// TIA Portal V20 export
Screen "OP01Pop-up_PRBWork"  274x350
  ScreenItem "Text field TG Status" at 1,0 size 273x47  Type=HmiTextBox
  ScreenItem "Cancel Mode" at 195,3 size 76x42  Type=HmiButton
  ScreenItem "Rectangle TG1" at 4,52 size 265x29  Type=HmiRectangle
  ScreenItem "Textfeld_1" at 9,57 size 21x20  Type=HmiTextBox
  ScreenItem "Textfeld_2" at 50,56 size 245x20  Type=HmiTextBox
  ScreenItem "Rectangle TG1_1" at 4,84 size 265x29  Type=HmiRectangle
  ScreenItem "Textfeld_5" at 9,88 size 21x20  Type=HmiTextBox
  ScreenItem "Rectangle TG1_2" at 4,116 size 265x29  Type=HmiRectangle
  ScreenItem "Textfeld_8" at 9,120 size 21x20  Type=HmiTextBox
  ScreenItem "Rectangle TG1_3" at 4,148 size 265x29  Type=HmiRectangle
  ScreenItem "Rectangle TG1_4" at 4,180 size 265x29  Type=HmiRectangle
  ScreenItem "Rectangle TG1_5" at 4,212 size 265x29  Type=HmiRectangle
  ScreenItem "Textfeld_3" at 50,88 size 245x20  Type=HmiTextBox
  ScreenItem "Textfeld_4" at 50,121 size 245x20  Type=HmiTextBox
  ScreenItem "Textfeld_7" at 50,153 size 245x20  Type=HmiTextBox
  ScreenItem "Textfeld_14" at 50,183 size 275x20  Type=HmiTextBox
  ScreenItem "Rectangle TG1_6" at 3,245 size 265x29  Type=HmiRectangle
  ScreenItem "Textfeld_6" at 9,151 size 21x20  Type=HmiTextBox
  ScreenItem "Textfeld_11" at 50,214 size 275x20  Type=HmiTextBox
  ScreenItem "Rectangle TG1_7" at 4,279 size 265x29  Type=HmiRectangle
  ScreenItem "Textfeld_10" at 9,185 size 21x20  Type=HmiTextBox
  ScreenItem "Rectangle TG1_8" at 4,314 size 265x29  Type=HmiRectangle
  ScreenItem "Textfeld_16" at 9,219 size 21x20  Type=HmiTextBox
  ScreenItem "Line_1" at 37,52 size 1x291  Type=HmiLine
  ScreenItem "Textfeld_9" at 52,250 size 275x20  Type=HmiTextBox
  ScreenItem "Textfeld_18" at 10,250 size 21x20  Type=HmiTextBox
